Yaskawa INFORM job: JUMPJOB.JBI

/JOB
//NAME JUMPJOB
//POS
///NPOS 1,0,0,0,0,0
///TOOL 0
///POSTYPE PULSE
///PULSE
C00000=-1,1,-2,-1,-64567,-1
//INST
///DATE 2025/10/28 03:33
///ATTR SC,RW
///GROUP1 RB1
NOP
MOVJ C00000 VJ=5.00
JUMP JOB:SQUIRCLE
END
